RoboDK station: demo-station.rdk

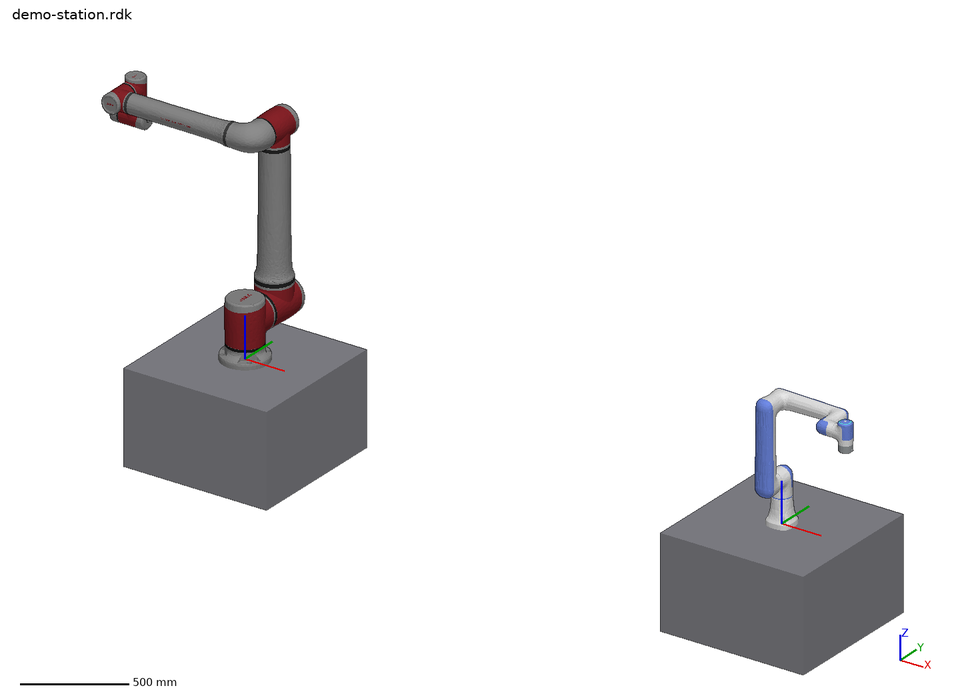
[picture v0: the station drawn from its stored meshes, robots at their saved joint values, targets as dots, program paths as lines]
Station demo-station (saved by RoboDK 5.9.0). Poses are relative to the parent item; angles as X-Y-Z fixed-axis rotations.
  - object Table JAKA at (0, 0, 0) mm, size 800 x 800 x 500 mm
  - frame JAKA Zu20 Base at (0, 0, 500) mm
    - robot JAKA Zu20: 6 axes
        modified DH rows (alpha deg, a mm, theta deg, d mm): 0, 0, 0, 196.5; 90, 0, 0, 0; 0, 897, 0, 0; 0, 744.5, 0, -188.35; 90, 0, 0, 138.5; -90, 0, 0, 120.5
        joint limits [-360, -85, -175, -85, -360, -360] to [360, 265, 175, 265, 360, 360]; home [0, 90, 90, 180, 90, 0]; saved at [0, 90, 90, 180, 90, 0]
  - object Table Nova 5 at (0, 0, 0) mm, size 800 x 800 x 500 mm
  - frame Dobot Nova 5 Base at (3000, 0, 500) mm
    - robot Dobot Nova 5: 6 axes
        modified DH rows (alpha deg, a mm, theta deg, d mm): 0, 0, 0, 240; 90, 0, 90, 0; 0, 400, 0, 0; 0, 330, -90, 135; -90, 0, 0, 120; 90, 0, 180, 88
        joint limits [-360, -180, -160, -360, -360, -360] to [360, 180, 160, 360, 360, 360]; home [0, 0, -90, 0, 90, 0]; saved at [0, 0, -90, 0, 90, 0]
